// TIA Portal V21 export
ORGANIZATION_BLOCK "Edges"   // OB1, LAD
   VAR_TEMP   // added for the SCL form of the ladder/FBD networks
      _w1 : Bool;
   END_VAR
BEGIN

REGION Network 1: Rising edge
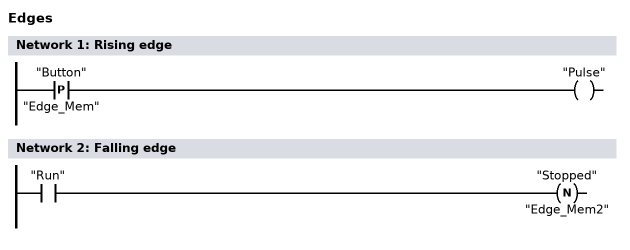
   #_w1 := "Button" AND NOT "Edge_Mem";   // rising edge of "Button"
   "Edge_Mem" := "Button";
   "Pulse" := #_w1;
END_REGION

REGION Network 2: Falling edge
   "Stopped" := NOT "Run" AND "Edge_Mem2";   // falling edge
   "Edge_Mem2" := "Run";
END_REGION
END_ORGANIZATION_BLOCK
